Staubli VAL3: placeInMatrix.pgx

program placeInMatrix(num nSlotIdx (byVal=true))
// Picks assembled unit from station and places it into the corresponding fMatrix slot.
  local num nRow
  local num nCol
  local point pCurPlace
  local point pCurApp
begin
  putln("[4/4] Placing assembly into matrix...")
  open(tLateral)

  // Pick assembled unit from assembling station
  movej(pAsmApproach, tLateral, mNomSpeed)
  waitEndMove()
  movel(pAsmCylinder, tLateral, mInsertSpeed)
  waitEndMove()
  close(tLateral)

  movel(pAsmApproach, tLateral, mNomSpeed)
  waitEndMove()

  // Compute (row, col) in 2x4 Assembled Matrix
  nRow = roundDown(nSlotIdx / nMatrixCols)
  nCol = nSlotIdx - (nRow * nMatrixCols)

  pCurPlace = pMatrixBase
  pCurPlace.trsf.x = pMatrixBase.trsf.x + (nCol * nMatrixStepX)
  pCurPlace.trsf.y = pMatrixBase.trsf.y + (nRow * nMatrixStepY)
  pCurApp = appro(pCurPlace, trMatrixAppro)

  putln("  -> Target matrix slot [" + toString("1.0", nRow) + "," + toString("1.0", nCol) + "]")

  movej(pCurApp, tLateral, mNomSpeed)
  waitEndMove()
  movel(pCurPlace, tLateral, mInsertSpeed)
  waitEndMove()
  open(tLateral)

  movel(pCurApp, tLateral, mNomSpeed)
  waitEndMove()
end
